Fanuc KAREL source: KA00186.KL

PROGRAM KA00186
%NOLOCKGROUP
VAR
  SRC: ARRAY[4] OF BYTE
  DST: ARRAY[4] OF SHORT
BEGIN
  DST = SRC
END KA00186
